SUBAPPLICATION SlurryTanker (* Subapplication Type *)
  (* Standard: 61499-2 *)
  (* Version 1.0, 2023-02-11, franz *)
  IMPORT DataPanel::io::MI::DQ::DataPanel_MI_DO::DigitalOutput_2A;
  IMPORT DataPanel::io::MI::DQ::DataPanel_MI_DO::DigitalOutput_2B;
  IMPORT DataPanel::io::MI::DQ::DataPanel_MI_DO::DigitalOutput_3A;
  IMPORT DataPanel::io::MI::DQ::DataPanel_MI_DO::DigitalOutput_3B;
  IMPORT DataPanel::io::MI::DQ::DataPanel_MI_DO::DigitalOutput_4A;
  IMPORT DataPanel::io::MI::DQ::DataPanel_MI_DO::DigitalOutput_4B;
  IMPORT DataPanel::io::MI::DQ::DataPanel_MI_DO::DigitalOutput_5A;
  IMPORT DataPanel::io::MI::DQ::DataPanel_MI_DO::DigitalOutput_5B;
  IMPORT DataPanel::io::MI::DQ::DataPanel_MI_DO::DigitalOutput_6A;
  IMPORT DataPanel::io::MI::DQ::DataPanel_MI_DO::DigitalOutput_7A;
  IMPORT DataPanel::io::MI::DQ::DataPanel_MI_DO::DigitalOutput_7B;
  IMPORT BlinkMarine::io::DI::PKP_2200_LI_DI::DigitalInput_Key_1;
  IMPORT BlinkMarine::io::DI::PKP_2200_LI_DI::DigitalInput_Key_2;
  IMPORT BlinkMarine::io::DI::PKP_2200_LI_DI::DigitalInput_Key_3;
  IMPORT BlinkMarine::io::DI::PKP_2200_LI_DI::DigitalInput_Key_4;
  IMPORT DefaultPool::AuxInput_Abscheider;
  IMPORT DefaultPool::AuxInput_Auseinanderklappen;
  IMPORT DefaultPool::AuxInput_Dom;
  IMPORT DefaultPool::AuxInput_Heckschieber;
  IMPORT DefaultPool::AuxInput_Knickdeichsel_heben;
  IMPORT DefaultPool::AuxInput_Knickdeichsel_senken;
  IMPORT DefaultPool::AuxInput_Licht;
  IMPORT DefaultPool::AuxInput_Schneidwerk;
  IMPORT DefaultPool::AuxInput_Seitenschieber;
  IMPORT DefaultPool::AuxInput_Verteiler_heben;
  IMPORT DefaultPool::AuxInput_Verteiler_senken;
  IMPORT DefaultPool::AuxInput_Zusammenklappen;
  IMPORT DefaultPool::SoftKey_Abscheider;
  IMPORT DefaultPool::SoftKey_Auseinanderklappen;
  IMPORT DefaultPool::SoftKey_Dom;
  IMPORT DefaultPool::SoftKey_Heckschieber;
  IMPORT DefaultPool::SoftKey_Knickdeichsel_heben;
  IMPORT DefaultPool::SoftKey_Knickdeichsel_senken;
  IMPORT DefaultPool::SoftKey_Licht;
  IMPORT DefaultPool::SoftKey_Schneidwerk;
  IMPORT DefaultPool::SoftKey_Seitenschieber;
  IMPORT DefaultPool::SoftKey_Verteiler_heben;
  IMPORT DefaultPool::SoftKey_Verteiler_senken;
  IMPORT DefaultPool::SoftKey_Zusammenklappen;
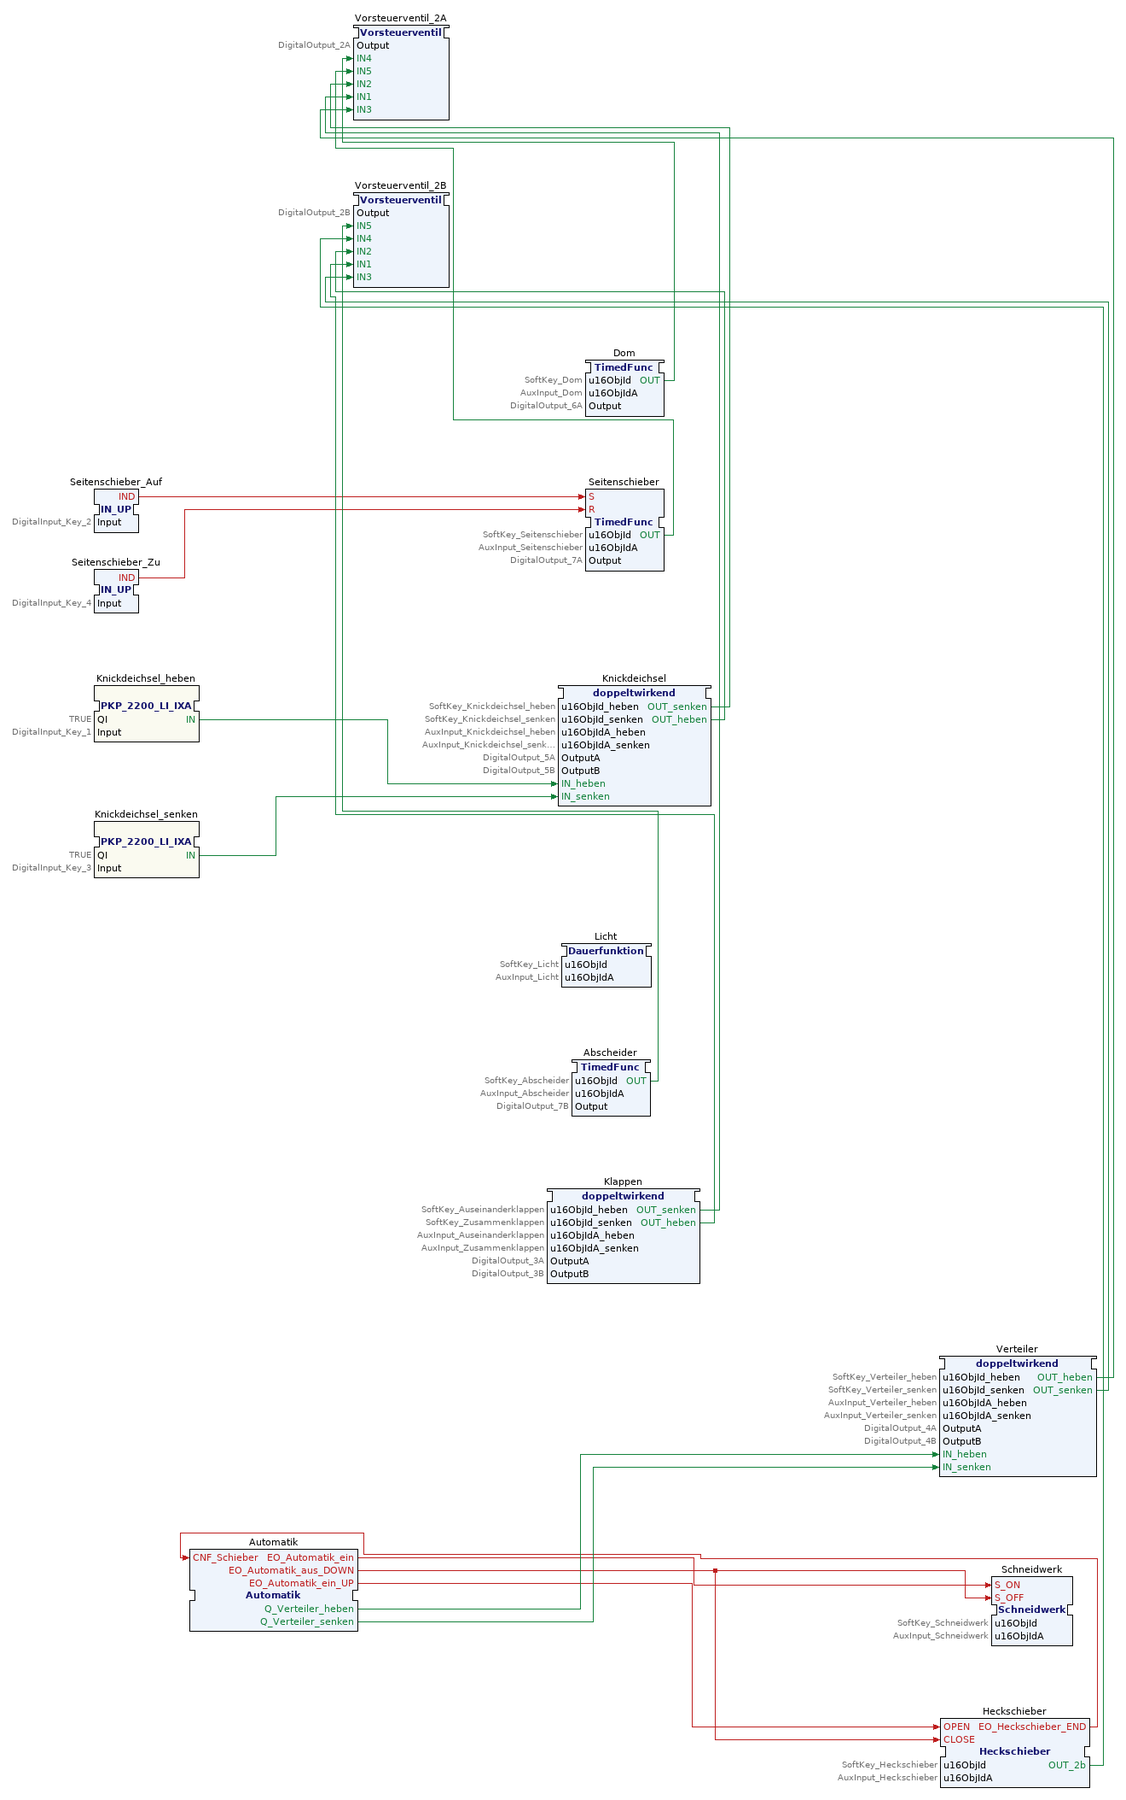
  (* Group funktionen: *)
  (* Group Vorsteuerventile: Vorsteuerventile *)
  (* Group Vorgewendeautomatik: Vorgewendeautomatik *)
  FBS
    Knickdeichsel_heben : BlinkMarine::io::DI::PKP_2200_LI_IXA(QI := TRUE, Input := DigitalInput_Key_1); {SET_ATTRIBUTE(GroupName, funktionen)}
    Knickdeichsel_senken : BlinkMarine::io::DI::PKP_2200_LI_IXA(QI := TRUE, Input := DigitalInput_Key_3); {SET_ATTRIBUTE(GroupName, funktionen)}
  END_FBS
  SUBAPPS
    Automatik : Automatik; {SET_ATTRIBUTE(GroupName, Vorgewendeautomatik)}
    Dom : TimedFunc(u16ObjId := SoftKey_Dom, u16ObjIdA := AuxInput_Dom, Output := DigitalOutput_6A); {SET_ATTRIBUTE(GroupName, funktionen)}
    Seitenschieber : TimedFunc(u16ObjId := SoftKey_Seitenschieber, u16ObjIdA := AuxInput_Seitenschieber, Output := DigitalOutput_7A); {SET_ATTRIBUTE(GroupName, funktionen)}
    Klappen : doppeltwirkend(u16ObjId_heben := SoftKey_Auseinanderklappen, u16ObjId_senken := SoftKey_Zusammenklappen, u16ObjIdA_heben := AuxInput_Auseinanderklappen, u16ObjIdA_senken := AuxInput_Zusammenklappen, OutputA := DigitalOutput_3A, OutputB := DigitalOutput_3B); {SET_ATTRIBUTE(GroupName, funktionen)}
    Verteiler : doppeltwirkend(u16ObjId_heben := SoftKey_Verteiler_heben, u16ObjId_senken := SoftKey_Verteiler_senken, u16ObjIdA_heben := AuxInput_Verteiler_heben, u16ObjIdA_senken := AuxInput_Verteiler_senken, OutputA := DigitalOutput_4A, OutputB := DigitalOutput_4B); {SET_ATTRIBUTE(GroupName, Vorgewendeautomatik)}
    Vorsteuerventil_2A : Vorsteuerventil(Output := DigitalOutput_2A); {SET_ATTRIBUTE(GroupName, Vorsteuerventile)}
    Vorsteuerventil_2B : Vorsteuerventil(Output := DigitalOutput_2B); {SET_ATTRIBUTE(GroupName, Vorsteuerventile)}
    Knickdeichsel : doppeltwirkend(u16ObjId_heben := SoftKey_Knickdeichsel_heben, u16ObjId_senken := SoftKey_Knickdeichsel_senken, u16ObjIdA_heben := AuxInput_Knickdeichsel_heben, u16ObjIdA_senken := AuxInput_Knickdeichsel_senken, OutputA := DigitalOutput_5A, OutputB := DigitalOutput_5B); {SET_ATTRIBUTE(GroupName, funktionen)}
    Licht : Dauerfunktion(u16ObjId := SoftKey_Licht, u16ObjIdA := AuxInput_Licht); {SET_ATTRIBUTE(GroupName, funktionen)}
    Abscheider : TimedFunc(u16ObjId := SoftKey_Abscheider, u16ObjIdA := AuxInput_Abscheider, Output := DigitalOutput_7B); {SET_ATTRIBUTE(GroupName, funktionen)}
    Schneidwerk : Schneidwerk(u16ObjId := SoftKey_Schneidwerk, u16ObjIdA := AuxInput_Schneidwerk); {SET_ATTRIBUTE(GroupName, Vorgewendeautomatik)}
    Heckschieber : Heckschieber(u16ObjId := SoftKey_Heckschieber, u16ObjIdA := AuxInput_Heckschieber); {SET_ATTRIBUTE(GroupName, Vorgewendeautomatik)}
    Seitenschieber_Auf : IN_UP(Input := DigitalInput_Key_2); {SET_ATTRIBUTE(GroupName, funktionen)}
    Seitenschieber_Zu : IN_UP(Input := DigitalInput_Key_4); {SET_ATTRIBUTE(GroupName, funktionen)}
  END_SUBAPPS
  EVENT_CONNECTIONS
    Automatik.EO_Automatik_ein TO Schneidwerk.S_ON;
    Automatik.EO_Automatik_aus_DOWN TO Schneidwerk.S_OFF;
    Automatik.EO_Automatik_ein_UP TO Heckschieber.OPEN;
    Automatik.EO_Automatik_aus_DOWN TO Heckschieber.CLOSE;
    Heckschieber.EO_Heckschieber_END TO Automatik.CNF_Schieber;
    Seitenschieber_Auf.IND TO Seitenschieber.S;
    Seitenschieber_Zu.IND TO Seitenschieber.R;
  END_CONNECTIONS
  ADAPTER_CONNECTIONS
    Dom.OUT TO Vorsteuerventil_2A.IN4;
    Seitenschieber.OUT TO Vorsteuerventil_2A.IN5;
    Abscheider.OUT TO Vorsteuerventil_2B.IN5;
    Heckschieber.OUT_2b TO Vorsteuerventil_2B.IN4;
    Automatik.Q_Verteiler_heben TO Verteiler.IN_heben;
    Automatik.Q_Verteiler_senken TO Verteiler.IN_senken;
    Knickdeichsel_heben.IN TO Knickdeichsel.IN_heben;
    Knickdeichsel_senken.IN TO Knickdeichsel.IN_senken;
    Knickdeichsel.OUT_senken TO Vorsteuerventil_2A.IN2;
    Knickdeichsel.OUT_heben TO Vorsteuerventil_2B.IN2;
    Klappen.OUT_senken TO Vorsteuerventil_2A.IN1;
    Klappen.OUT_heben TO Vorsteuerventil_2B.IN1;
    Verteiler.OUT_heben TO Vorsteuerventil_2A.IN3;
    Verteiler.OUT_senken TO Vorsteuerventil_2B.IN3;
  END_CONNECTIONS
END_SUBAPPLICATION
